(* IEC 61131-3 sources: Test-Git_ESME26/TestProgettoESME_26.fbsproj/PacDriveLib Migration/Motion/Positioning/PDL_FB_EndlessFeed.fb.st^, 8 files *)

(* ---- Init.meth.st ---- *)
METHOD PRIVATE Init : BOOL
VAR_INPUT
END_VAR

Init := FALSE;

IF i_ifDrive = 0 THEN
	SetDiagOutput(	i_etDiag	:= GD.ET_Diag.InputParameterInvalid,
					i_etDiagExt := PDL_ET_DiagExt.DriveInvalid,
					i_sMsg		:= 'i_ifDrive - Invalid Interface');
	RETURN;

ELSIF NOT i_ifDrive.xIsHomed  THEN
	SetDiagOutput(	i_etDiag	:= GD.ET_Diag.DriveConditionInvalid,
					i_etDiagExt := PDL_ET_DiagExt.DriveNotHomed,
					i_sMsg		:= 'i_ifDrive - must be homed');
	RETURN;

ELSE
	//get IF_DriveConfig
	xSuccess := __QUERYINTERFACE(i_ifDrive, ifGetParentDevice);
	IF xSuccess AND ifGetParentDevice <> 0 THEN
		ifDeviceAccess := ifGetParentDevice.GetParentDevice();
		xSuccess := __QUERYINTERFACE( ifDeviceAccess, ifDriveConfigAccess );
		IF xSuccess AND ifDriveConfigAccess <> 0 THEN
			ifDriveConfig := ifDriveConfigAccess.DriveConfig;
		END_IF
	END_IF

	xSuccess := __QUERYINTERFACE(ifDeviceAccess, ifDeviceTreeObjectAccess);
	IF xSuccess THEN
		sDriveName := ifDeviceTreeObjectAccess.DeviceTreeObject.Name;
	ELSE
		sDriveName := 'Axis';
	END_IF

	fbStop.Axis := i_ifDrive;
	fbHalt.Axis := i_ifDrive;
	fbMoveAbsolute.Axis := i_ifDrive;
	fbMoveVelocity.Axis := i_ifDrive;

	//check axis
	xModuloAxis := i_ifDrive.xIsModulo;
	IF xModuloAxis THEN
		lrModuloPeriod 	:= i_ifDrive.lrModuloPeriod;
	END_IF
END_IF

Init := TRUE;

(* ---- InputParameterCheck.meth.st ---- *)
METHOD PRIVATE InputParameterCheck : BOOL
VAR_INPUT
END_VAR
VAR
	lrMaxAcc	: LREAL := 0;
	lrMaxVel	: LREAL := 0;
END_VAR

InputParameterCheck := FALSE;

//if IF_DriveConfig is not available -> limits are NOT checked
IF ifDriveConfig <> 0 THEN
	lrMaxAcc := ifDriveConfig.MaxAcc;
	lrMaxVel := ifDriveConfig.MaxVel;
END_IF

IF    NOT xModuloAxis
  AND i_lrPeriod <= 0.0
THEN
	SetDiagOutput(	i_etDiag	:= GD.ET_Diag.InputParameterInvalid,
					i_etDiagExt := PDL_ET_DiagExt.PeriodRange,
					i_sMsg		:= '0.0 < i_lrPeriod');

ELSIF i_lrStopPosition < 0.0 THEN
	SetDiagOutput(	i_etDiag	:= GD.ET_Diag.InputParameterInvalid,
					i_etDiagExt := PDL_ET_DiagExt.StopPositionRange,
					i_sMsg		:= '0.0 <= i_lrStopPosition');

ELSIF    xModuloAxis
	 AND i_lrStopPosition > lrModuloPeriod
THEN
	SetDiagOutput(	i_etDiag	:= GD.ET_Diag.InputParameterInvalid,
					i_etDiagExt := PDL_ET_DiagExt.StopPositionRange,
					i_sMsg		:= 'i_lrStopPosition > Modulo Period');

ELSIF i_lrAcc <= 0.0 OR (i_lrAcc > lrMaxAcc AND lrMaxAcc <> 0) THEN
	SetDiagOutput(	i_etDiag	:= GD.ET_Diag.InputParameterInvalid,
					i_etDiagExt := PDL_ET_DiagExt.AccRange,
					i_sMsg		:= STANDARD.CONCAT('0.0 < i_lrAcc <= ', TO_STRING(lrMaxAcc) ));

ELSIF i_lrDec <= 0.0 OR (i_lrDec > lrMaxAcc AND lrMaxAcc <> 0) THEN
	SetDiagOutput(	i_etDiag	:= GD.ET_Diag.InputParameterInvalid,
					i_etDiagExt := PDL_ET_DiagExt.DecRange,
					i_sMsg		:= STANDARD.CONCAT('0.0 < i_lrDec <= ', TO_STRING(lrMaxAcc) ));

ELSIF ABS(i_lrVel) > lrMaxVel AND lrMaxVel <> 0 THEN
	SetDiagOutput(	i_etDiag	:= GD.ET_Diag.InputParameterInvalid,
					i_etDiagExt := PDL_ET_DiagExt.VelRange,
					i_sMsg		:= STANDARD.CONCAT('0.0 < i_lrVel <= ', TO_STRING(lrMaxVel) ));

ELSIF i_lrJerk <= 0.0  THEN
	SetDiagOutput(	i_etDiag	:= GD.ET_Diag.InputParameterInvalid,
					i_etDiagExt := PDL_ET_DiagExt.JerkRange,
					i_sMsg		:= '0.0 < i_lrJerk');

ELSE
	InputParameterCheck := TRUE;
END_IF

(* ---- MoveToStopPosition.meth.st ---- *)
METHOD PRIVATE MoveToStopPosition : BOOL
VAR
	lrStopPosCycles      : LREAL;
	lrNormalizedStopPos  : LREAL;
	lrBrakePosCycles     : LREAL;
	lrNormalizedBrakePos : LREAL;
END_VAR

IF NOT InputParameterCheck() THEN

	q_xInVelocity				:= FALSE;
	q_xMotionInstructionActive	:= FALSE;
	q_xReady					:= FALSE;

	diState := 100;
ELSE
	q_xMotionInstructionActive := TRUE;

	// if velocity was set to zero together with i_xStart = FALSE take velocity of last seen command.
	IF i_lrVel <> 0 THEN
		lrActVel	:= i_lrVel;
	END_IF
	lrActJerk	:= i_lrJerk;
	lrAccel	:= i_lrACC;
	lrDecel	:= i_lrDEC;

	//calc new stop position
	IF NOT xMoveToStoppingStarted THEN

		//modulo axis
		IF xModuloAxis THEN
			lrStopPosition := i_lrStopPosition;

		//linear axis -> lrStopPosition has to be calculated
		ELSE
			IF lrActVel >= 0 THEN
				etResultCalcStopping := MOIN.FC_CalculateMoveVelocity( 	i_etDirection 				:= MOIN.ET_Direction.PositiveDirection, //not considered when TargetVelocity = 0
																		i_lrStartVelocity			:= i_ifDrive.lrVelocity + i_ifDrive.lrAcceleration*0.01,//tolerance to avoid overshoot
																		i_lrStartAcceleration		:= i_ifDrive.lrAcceleration,
																		i_lrMovementAcceleration 	:= lrAccel,
																		i_lrMovementDeceleration	:= lrDecel,
																		i_lrJerk 					:= lrActJerk,
																		i_lrStartPosition			:= 0.0, //inside a distance is calculated, StartPosition is added
																		i_lrTargetVelocity			:= 0.0,
																		q_stTrajectory				=> stStoppingDistance,
																		q_xError					=> xErrorCalcStopping
																		);
				IF xErrorCalcStopping THEN
					q_xActive					:= FALSE;
					q_xMotionInstructionActive	:= FALSE;
					q_lrPosition				:= 0.0;

					SetDiagOutput(	i_etDiag	:= GD.ET_Diag.UnexpectedProgramBehavior,
									i_etDiagExt := PDL_ET_DiagExt.UnexpectedFeedback,
									i_sMsg		:= CONCAT('FC_CalculateMoveVelocity.ET_Result: ', MOIN.FC_EtResultToString(etResultCalcStopping) ));
					diState := 100;
					RETURN;
				ELSE
					lrStoppingDistance := ABS(stStoppingDistance.astPoints[stStoppingDistance.uiNumberOfPhases].lrPosition);
				END_IF

				IF i_lrPeriod > 0 THEN
					lrPeriodeCount := DINT_TO_LREAL(TRUNC((q_lrPosition + lrStoppingDistance) / i_lrPeriod));
					IF q_lrPosition + lrStoppingDistance - lrPeriodeCount * i_lrPeriod > i_lrStopPosition THEN
						lrPeriodeCount := lrPeriodeCount + 1;
					END_IF
					lrStopPosition := i_lrStopPosition + lrPeriodeCount * i_lrPeriod;
				ELSE
					lrStopPosition := i_lrStopPosition;
				END_IF

			ELSE
				etResultCalcStopping := MOIN.FC_CalculateMoveVelocity( 	i_etDirection 				:= MOIN.ET_Direction.NegativeDirection,  //not considered when TargetVelocity = 0
																		i_lrStartVelocity			:= i_ifDrive.lrVelocity + i_ifDrive.lrAcceleration*0.01,//tolerance to avoid overshoot
																		i_lrStartAcceleration		:= i_ifDrive.lrAcceleration,
																		i_lrMovementAcceleration 	:= lrAccel,
																		i_lrMovementDeceleration	:= lrDecel,
																		i_lrJerk 					:= lrActJerk,
																		i_lrStartPosition			:= 0,
																		i_lrTargetVelocity			:= 0.0,
																		q_stTrajectory				=> stStoppingDistance,
																		q_xError					=> xErrorCalcStopping
																		);
				IF xErrorCalcStopping THEN
					q_xActive					:= FALSE;
					q_xMotionInstructionActive	:= FALSE;
					q_lrPosition				:= 0.0;

					SetDiagOutput(	i_etDiag	:= GD.ET_Diag.UnexpectedProgramBehavior,
									i_etDiagExt := PDL_ET_DiagExt.UnexpectedFeedback,
									i_sMsg		:= CONCAT('FC_CalculateMoveVelocity.ET_Result: ', MOIN.FC_EtResultToString(etResultCalcStopping) ));
					diState := 100;
					RETURN;
				ELSE
					lrStoppingDistance := ABS(stStoppingDistance.astPoints[stStoppingDistance.uiNumberOfPhases].lrPosition);
				END_IF

				IF i_lrPeriod > 0 THEN
					lrStopPosCycles      := TO_LREAL(TRUNC(i_lrStopPosition / i_lrPeriod));
					lrNormalizedStopPos  := i_lrStopPosition - lrStopPosCycles * i_lrPeriod;
					lrBrakePosCycles     := ABS(TO_LREAL(TRUNC((q_lrPosition - lrStoppingDistance - i_lrPeriod) / i_lrPeriod))); // slided one period to negative, because first negative period would be zero (as "first" positive period)
					lrNormalizedBrakePos := q_lrPosition - lrStoppingDistance + lrBrakePosCycles * i_lrPeriod;
					IF lrStopPosCycles >= 1.0 OR lrNormalizedBrakePos > lrNormalizedStopPos THEN
						// can stop in cycle or is forced to move to next cycle with too big i_lrStopPosition anyway
						lrStopPosition := lrNormalizedStopPos - (lrStopPosCycles + lrBrakePosCycles) * i_lrPeriod;
					ELSE
						// add additional move to next cycle to prevent overswing
						lrStopPosition := lrNormalizedStopPos - (lrStopPosCycles + lrBrakePosCycles + 1.0) * i_lrPeriod;
					END_IF
				ELSE
					lrStopPosition := i_lrStopPosition;
				END_IF
			END_IF
		END_IF
	END_IF

	//reset fbs
	fbMoveVelocity( Execute := FALSE);
	fbMoveAbsolute( Execute := FALSE);

	//call fb with new values
	fbMoveAbsolute(	Execute			:= TRUE,
					Position		:= lrStopPosition,
					Velocity		:= ABS(lrActVel),
					Acceleration	:= lrAccel,
					Deceleration	:= lrDecel,
					Jerk			:= lrActJerk,
					Direction		:= fbMoveVelocity.Direction);

	//set output msg
	SetDiagOutput(	i_etDiag	:= GD.ET_Diag.Ok,
					i_etDiagExt := PDL_ET_DiagExt.WaitUntilStopPositionReached,
					i_sMsg		:= '');

END_IF

(* ---- MoveVelocity.meth.st ---- *)
METHOD PRIVATE MoveVelocity : BOOL
VAR_INPUT
END_VAR

IF NOT InputParameterCheck() THEN

	q_xInVelocity				:= FALSE;
	q_xMotionInstructionActive	:= FALSE;
	q_xReady					:= FALSE;

	diState := 100;
ELSE
	q_xMotionInstructionActive := TRUE;

	//check if velocity changes direction
	IF (lrActVel*i_lrVel) >= 0 THEN
		lrAccel	:= i_lrACC;
		lrDecel	:= i_lrDEC;
	ELSE //if yes take acceleration also for deceleration phase
		lrAccel	:= i_lrACC;
		lrDecel	:= i_lrACC;
	END_IF
	lrActVel  := i_lrVel;
	lrActJerk := i_lrJerk;

	//set direction
	IF lrActVel < 0 THEN
		fbMoveVelocity.Direction := MOIN.ET_Direction.NegativeDirection;
	ELSE
		fbMoveVelocity.Direction := MOIN.ET_Direction.PositiveDirection;
	END_IF

	//reset fbs
	fbMoveAbsolute( Execute := FALSE);
	fbMoveVelocity( Execute := FALSE );

	//call fb with new values
	fbMoveVelocity(	Execute			:= TRUE,
					Velocity		:= ABS(lrActVel),
					Acceleration	:= lrAccel,
					Deceleration	:= lrDecel,
					Jerk			:= lrActJerk);

	//set output msg
	SetDiagOutput(	i_etDiag	:= GD.ET_Diag.Ok,
					i_etDiagExt := PDL_ET_DiagExt.EndlessPositioning,
					i_sMsg		:= Standard.CONCAT('Velocity: ', LREAL_TO_STRING(lrActVel)));

END_IF

(* ---- RegisterLoggerPoint.meth.st ---- *)
METHOD PUBLIC RegisterLoggerPoint
VAR_INPUT
	i_ifParent		: APL.IF_LoggerPoint;
	i_sName			: STRING[80];
END_VAR
VAR_OUTPUT
	q_etDiag		: GD.ET_Diag := GD.ET_Diag.Ok;
	q_etDiagExt		: PDL_ET_DiagExt := PDL_ET_DiagExt.Ok;
END_VAR
VAR
	etDiagBuffer		: GD.ET_Diag;
	etDiagExtBufferAPL	: APL.ET_DiagExt;
END_VAR

fbLoggerPoint.RegisterLoggerPoint(	i_ifParent		:= i_ifParent,
									i_sName			:= i_sName,
									i_sType			:= 'FB_EndlessFeed',
									i_sSource		:= 'PDL',
									q_etDiag		=> etDiagBuffer,
									q_etDiagExt		=> etDiagExtBufferAPL);
IF (etDiagBuffer <> GD.ET_Diag.Ok) THEN
	CASE etDiagExtBufferAPL OF
		APL.ET_DiagExt.ParentInvalid:
			q_etDiag := GD.ET_Diag.InputParameterInvalid;
			q_etDiagExt := PDL_ET_DiagExt.ParentInvalid;

		APL.ET_DiagExt.ParentNotRegistered:
			q_etDiag := GD.ET_Diag.InputParameterInvalid;
			q_etDiagExt := PDL_ET_DiagExt.ParentNotRegistered;

		APL.ET_DiagExt.MaxNumberOfLoggerPointsExeeded:
			q_etDiag := GD.ET_Diag.InputParameterInvalid;
			q_etDiagExt := PDL_ET_DiagExt.MaxNumberOfLoggerPointsExeeded;

	ELSE
		q_etDiag := GD.ET_Diag.UnexpectedProgramBehavior;
		q_etdiagExt := PDL_ET_DiagExt.UnexpectedDiagExt;
	END_CASE
END_IF

(* ---- SetDiagOutput.meth.st ---- *)
METHOD PRIVATE SetDiagOutput : BOOL
VAR_INPUT
	i_etDiag	: GD.ET_Diag;
	i_etDiagExt	: PDL_ET_DiagExt;
	i_sMsg		: STRING[80];
END_VAR
VAR
END_VAR

IF i_etDiag <> GD.ET_Diag.Ok THEN
	q_xReady := FALSE;
END_IF
IF q_etDiag = GD.ET_Diag.OK OR i_etDiagExt = PDL_ET_DiagExt.Disabled THEN
	q_etDiag := i_etDiag;
	q_etDiagExt := i_etDiagExt;
	q_sMsg := i_sMsg;

	IF(i_etDiag = GD.ET_Diag.Ok) AND (fbLoggerPoint.etLogLevel >= APL.ET_LogLevel.StatusMessage) THEN
		fbLoggerPoint.AddLogEntry(	i_etLogLevel	:= APL.ET_LogLevel.StatusMessage,
									i_etDiag		:= q_etDiag,
									i_udiDiagExt	:= q_etDiagExt,
									i_sMessage		:= SE_CTBX.FC_MultiConcat(	i_sString1	:= Standard.CONCAT('ET_Diag: ', GD.FC_EtDiagToString(q_etDiag)),
																				i_sString2	:= Standard.CONCAT(' ET_DiagExt: ', PDL_FC_EtDiagExtToString(q_etDiagExt)),
																				i_sString3	:= Standard.CONCAT(' sMsg: ', q_sMsg),
																				i_sString4	:= '')
									);
	ELSIF(i_etDiag = GD.ET_Diag.UnexpectedProgramBehavior) AND (fbLoggerPoint.etLogLevel >= APL.ET_LogLevel.CriticalException) THEN
		fbLoggerPoint.AddLogEntry(	i_etLogLevel	:= APL.ET_LogLevel.CriticalException,
									i_etDiag		:= q_etDiag,
									i_udiDiagExt	:= q_etDiagExt,
									i_sMessage		:= SE_CTBX.FC_MultiConcat(	i_sString1	:= Standard.CONCAT('ET_Diag: ', GD.FC_EtDiagToString(q_etDiag)),
																				i_sString2	:= Standard.CONCAT(' ET_DiagExt: ', PDL_FC_EtDiagExtToString(q_etDiagExt)),
																				i_sString3	:= Standard.CONCAT(' sMsg: ', q_sMsg),
																				i_sString4	:= '')
									);
	ELSIF(i_etDiag <> GD.ET_Diag.Ok) AND (fbLoggerPoint.etLogLevel >= APL.ET_LogLevel.Exception) THEN
		fbLoggerPoint.AddLogEntry(	i_etLogLevel	:= APL.ET_LogLevel.Exception,
									i_etDiag		:= q_etDiag,
									i_udiDiagExt	:= q_etDiagExt,
									i_sMessage		:= SE_CTBX.FC_MultiConcat(	i_sString1	:= Standard.CONCAT('ET_Diag: ', GD.FC_EtDiagToString(q_etDiag)),
																				i_sString2	:= Standard.CONCAT(' ET_DiagExt: ', PDL_FC_EtDiagExtToString(q_etDiagExt)),
																				i_sString3	:= Standard.CONCAT(' sMsg: ', q_sMsg),
																				i_sString4	:= '')
									);
	END_IF
END_IF

(* ---- SetInVelocity.meth.st ---- *)
METHOD PRIVATE SetInVelocity : BOOL
VAR_INPUT
END_VAR
VAR
	lrMaxVelDeviation			: LREAL;
	lrCurrVelDeviation			: LREAL;
END_VAR

// Check, if we have already reached the required velocity
IF (ABS(lrActVel) > 0) THEN

	lrMaxVelDeviation	:= 0.01 * ABS(i_ifDrive.lrVelocity);
	lrCurrVelDeviation	:= ABS( lrActVel - i_ifDrive.lrVelocity);
	IF (lrCurrVelDeviation <= lrMaxVelDeviation )THEN
		q_xInVelocity	:= TRUE;
	ELSE
		q_xInVelocity	:= FALSE;
	END_IF
ELSE
	q_xInVelocity := q_xMotionInstructionActive;
END_IF

(* ---- SetPos.meth.st ---- *)
METHOD PRIVATE SetPos : BOOL
VAR_INPUT
END_VAR

IF i_lrPeriod > 0 THEN

	//reset fb
	fbSetPos(	Axis := i_ifDrive, Execute := FALSE );

	IF (q_lrPosition > 2 * i_lrPeriod) OR q_lrPosition  < -i_lrPeriod THEN
		lrPeriodeCount := TRUNC_INT(q_lrPosition / i_lrPeriod);
		IF q_lrPosition < 0 THEN
			lrPeriodeCount := (lrPeriodeCount - 1);
		END_IF

		IF lrPeriodeCount <> 0 THEN
			q_lrPosition:= q_lrPosition - lrPeriodeCount * i_lrPeriod;

			fbSetPos(	Axis		:= i_ifDrive,
						Execute		:= TRUE,
						Position	:= -lrPeriodeCount * i_lrPeriod,
						Relative	:= TRUE);

			IF fbSetPos.Error THEN
				SetDiagOutput(	i_etDiag	:= GD.ET_Diag.UnexpectedProgramBehavior,
								i_etDiagExt := PDL_ET_DiagExt.UnexpectedFeedback,
								i_sMsg		:= CONCAT('MC_SetPosition.ErrorId: ', TO_STRING(fbSetPos.ErrorId)));
				RETURN;
			END_IF

			lrStopPosition := lrStopPosition - lrPeriodeCount * i_lrPeriod;
		END_IF

	ELSIF q_lrPosition > i_lrPeriod + 0.001  THEN
		lrInchPos		:= lrInchPos - i_lrPeriod;
		q_lrPosition	:= q_lrPosition - i_lrPeriod;

		fbSetPos(	Axis		:= i_ifDrive,
					Execute		:= TRUE,
					Position	:= -i_lrPeriod,
					Relative	:= TRUE);

		IF fbSetPos.Error THEN
			SetDiagOutput(	i_etDiag	:= GD.ET_Diag.UnexpectedProgramBehavior,
							i_etDiagExt := PDL_ET_DiagExt.UnexpectedFeedback,
							i_sMsg		:= CONCAT('MC_SetPosition.ErrorId: ', TO_STRING(fbSetPos.ErrorId)));
			RETURN;
		END_IF

		lrStopPosition := lrStopPosition - i_lrPeriod;

	ELSIF q_lrPosition  < -0.001 THEN
		lrInchPos		:= lrInchPos + i_lrPeriod;
		q_lrPosition	:= q_lrPosition + i_lrPeriod;

		fbSetPos(	Axis		:= i_ifDrive,
					Execute		:= TRUE,
					Position	:= i_lrPeriod,
					Relative	:= TRUE);

		IF fbSetPos.Error THEN
			SetDiagOutput(	i_etDiag	:= GD.ET_Diag.UnexpectedProgramBehavior,
							i_etDiagExt := PDL_ET_DiagExt.UnexpectedFeedback,
							i_sMsg		:= CONCAT('MC_SetPosition.ErrorId: ', TO_STRING(fbSetPos.ErrorId)));
			RETURN;
		END_IF

		lrStopPosition := lrStopPosition + i_lrPeriod;
	END_IF
END_IF
